TYPE ST_PIDOperatorValues :
STRUCT
	setpoint			: LREAL; //operator setpoint in PV units (Setpoint mode)
	ratio				: LREAL; //operator ratio (Ratio mode)
	output				: LREAL; //operator output in % (OpenLoop mode)
END_STRUCT
END_TYPE

(* stored: Version 1.1.0.1, ProductVersion 3.1.4024.12
   DUT ST_PIDOperatorValues: Id {3bc1dea2-5e7e-4a92-b3fd-94c81c13fd14} *)
